Staubli VAL3: moveTarget.pgx

public program moveTarget(point x_pTarget, joint x_jTarget)
  local bool l_bEqual
  local joint l_jCurrentPosUp
  local joint l_jTargetPosUp
  local point l_pCurrentPosUp
  local point l_pTargetPosUp
  local bool l_bOK1
  local bool l_bOK2
  local num l_nDir
begin
  switch sMounting
    case "Floor"
      l_nDir=1
    break
    case "Ceiling"
      l_nDir=-1
    break
    default
      l_nDir=1
    break
  endSwitch
  //
  call CheckPosEqual(x_pTarget,l_bEqual)
  if l_bEqual==false
    call hmiAlert("Move","info")
    l_pCurrentPosUp=compose(here(utCurrentTool.tValue,world),world,{0,0,100*l_nDir,0,0,0})
    l_bOK1=pointToJoint(utCurrentTool.tValue,x_jTarget,l_pCurrentPosUp,l_jCurrentPosUp)
    l_pTargetPosUp=compose(x_pTarget,world,{0,0,100*l_nDir,0,0,0})
    l_bOK2=pointToJoint(utCurrentTool.tValue,x_jTarget,l_pTargetPosUp,l_jTargetPosUp)
    if l_bOK1==true and l_bOK2==true
      movel(l_pCurrentPosUp,utCurrentTool.tValue,mSpeed_J_blend)
      movej(l_jTargetPosUp,utCurrentTool.tValue,mSpeed_J_blend)
      movel(compose(x_pTarget,world,{0,0,20*l_nDir,0,0,0}),utCurrentTool.tValue,mSpeed_J_blend)
      movel(x_pTarget,utCurrentTool.tValue,mSlow)
      waitEndMove()
      call hmiAlert("CompleteMove","info")
    else
      call hmiAlert("CantMove2","warning")
    endIf
  else
    call hmiAlert("CompleteMove","info")
  endIf
end
